// TIA Portal V17 export
// export: Created 2000-01-01T00:00:00.0000000Z, ExportSetting None
FUNCTION "FC_Rung" : Void   // FC42, LAD
{ S7_Optimized_Access := 'TRUE' }
   VAR_INPUT
      Local : Int;
   END_VAR
BEGIN

REGION Network 1
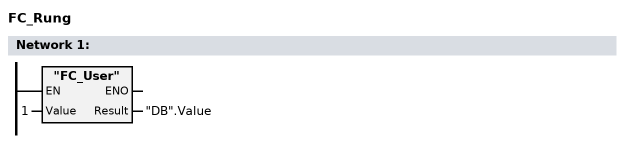
   RUNG wire#powerrail
      "FC_User"(Value := 1, Result => "DB".Value)
   END_RUNG
   // the same network as SCL:
   "FC_User"(Value := 1, Result => "DB".Value);
END_REGION
END_FUNCTION
